Fanuc KAREL source: KT00684.KL

PROGRAM KT00684
%NOLOCKGROUP
VAR
  P1: JOINTPOS
  P2: JOINTPOS
  OUT: BOOLEAN
BEGIN
  OUT = + P1
END KT00684
